// TIA Portal V19 export
DATA_BLOCK "CV_DATA"   // DB17
{ S7_Optimized_Access := 'FALSE' }
   VAR
      CHILLED_SKID_P01 : Struct
         CMD : Bool;
         SET_POINT : Real;
         INPUT : Real;
         OUT_PUT : Real;
         OUTPUT_PER : Int;
         NORM_MIN : Int;
         NORM_MAX : Int := 27684;
         NORM_OUT : Real;
         SCALE_MIN : Real;
         SCALE_MAX : Real := 50.0;
         SCALE_OUT : Real;
         MANUAL_OPEN_PER : Int;
         MANUAL_TEMP : Int;
         MANOUT : Real;
         PUMP_AO : Real;
      END_STRUCT;
      HS_PCV801 : Struct
         CMD : Bool;
         SET_POINT : Real;
         INPUT : Real;
         OUT_PUT : Real;
         OUTPUT_PER : Int;
         NORM_MIN : Int;
         NORM_MAX : Int;
         NORM_OUT : Real;
         SCALE_MIN : Real;
         SCALE_MAX : Real;
         SCALE_OUT : Real;
         MANUAL_OPEN_PER : Int;
         MANUAL_TEMP : Int;
         MANOUT : Int;
         CV_AO : Int;
      END_STRUCT;
      CHILLED_SKID_P02 : Struct
         CMD : Bool;
         SET_POINT : Real;
         INPUT : Real;
         OUT_PUT : Real;
         OUTPUT_PER : Int;
         NORM_MIN : Int;
         NORM_MAX : Int := 27684;
         NORM_OUT : Real := 0.0;
         SCALE_MIN : Real := 0.0;
         SCALE_MAX : Real := 50.0;
         SCALE_OUT : Real;
         MANUAL_OPEN_PER : Int;
         MANUAL_TEMP : Int;
         MANOUT : Real;
         PUMP_AO : Real;
      END_STRUCT;
      CHILLED_SKID_P03 : Struct
         CMD : Bool;
         SET_POINT : Real;
         INPUT : Real;
         OUT_PUT : Real;
         OUTPUT_PER : Int;
         NORM_MIN : Int;
         NORM_MAX : Int := 27684;
         NORM_OUT : Real := 0.0;
         SCALE_MIN : Real := 0.0;
         SCALE_MAX : Real := 50.0;
         SCALE_OUT : Real;
         MANUAL_OPEN_PER : Int;
         MANUAL_TEMP : Int;
         MANOUT : Real;
         PUMP_AO : Real;
      END_STRUCT;
      HOT_SKID_P01 : Struct
         CMD : Bool;
         SET_POINT : Real;
         INPUT : Real;
         OUT_PUT : Real;
         OUTPUT_PER : Int;
         NORM_MIN : Int;
         NORM_MAX : Int := 27684;
         NORM_OUT : Real := 0.0;
         SCALE_MIN : Real := 0.0;
         SCALE_MAX : Real := 50.0;
         SCALE_OUT : Real;
         MANUAL_OPEN_PER : Int;
         MANUAL_TEMP : Int;
         MANOUT : Real;
         PUMP_AO : Real;
      END_STRUCT;
      HOT_SKID_P02 : Struct
         CMD : Bool;
         SET_POINT : Real;
         INPUT : Real;
         OUT_PUT : Real;
         OUTPUT_PER : Int;
         NORM_MIN : Int;
         NORM_MAX : Int := 27684;
         NORM_OUT : Real := 0.0;
         SCALE_MIN : Real := 0.0;
         SCALE_MAX : Real := 50.0;
         SCALE_OUT : Real;
         MANUAL_OPEN_PER : Int;
         MANUAL_TEMP : Int;
         MANOUT : Real;
         PUMP_AO : Real;
      END_STRUCT;
      HOT_SKID_P03 : Struct
         CMD : Bool;
         SET_POINT : Real;
         INPUT : Real;
         OUT_PUT : Real;
         OUTPUT_PER : Int;
         NORM_MIN : Int;
         NORM_MAX : Int := 27684;
         NORM_OUT : Real := 0.0;
         SCALE_MIN : Real := 0.0;
         SCALE_MAX : Real := 50.0;
         SCALE_OUT : Real;
         MANUAL_OPEN_PER : Int;
         MANUAL_TEMP : Int;
         MANOUT : Real;
         PUMP_AO : Real;
      END_STRUCT;
      COLD_SKID_P01 : Struct
         CMD : Bool;
         SET_POINT : Real;
         INPUT : Real;
         OUT_PUT : Real;
         OUTPUT_PER : Int;
         NORM_MIN : Int;
         NORM_MAX : Int := 27684;
         NORM_OUT : Real := 0.0;
         SCALE_MIN : Real := 0.0;
         SCALE_MAX : Real := 50.0;
         SCALE_OUT : Real;
         MANUAL_OPEN_PER : Int;
         MANUAL_TEMP : Int;
         MANOUT : Real;
         PUMP_AO : Real;
      END_STRUCT;
      COLD_SKID_P02 : Struct
         CMD : Bool;
         SET_POINT : Real;
         INPUT : Real;
         OUT_PUT : Real;
         OUTPUT_PER : Int;
         NORM_MIN : Int;
         NORM_MAX : Int := 27684;
         NORM_OUT : Real := 0.0;
         SCALE_MIN : Real := 0.0;
         SCALE_MAX : Real := 50.0;
         SCALE_OUT : Real;
         MANUAL_OPEN_PER : Int;
         MANUAL_TEMP : Int;
         MANOUT : Real;
         PUMP_AO : Real;
      END_STRUCT;
      COLD_SKID_P03 : Struct
         CMD : Bool;
         SET_POINT : Real;
         INPUT : Real;
         OUT_PUT : Real;
         OUTPUT_PER : Int;
         NORM_MIN : Int;
         NORM_MAX : Int := 27684;
         NORM_OUT : Real := 0.0;
         SCALE_MIN : Real := 0.0;
         SCALE_MAX : Real := 50.0;
         SCALE_OUT : Real;
         MANUAL_OPEN_PER : Int;
         MANUAL_TEMP : Int;
         MANOUT : Real;
         PUMP_AO : Real;
      END_STRUCT;
      UCH_SKID_P01 : Struct
         CMD : Bool;
         SET_POINT : Real;
         INPUT : Real;
         OUT_PUT : Real;
         OUTPUT_PER : Int;
         NORM_MIN : Int;
         NORM_MAX : Int := 27684;
         NORM_OUT : Real := 0.0;
         SCALE_MIN : Real := 0.0;
         SCALE_MAX : Real := 50.0;
         SCALE_OUT : Real;
         MANUAL_OPEN_PER : Int;
         MANUAL_TEMP : Int;
         MANOUT : Real;
         PUMP_AO : Real;
      END_STRUCT;
      UCH_SKID_P02 : Struct
         CMD : Bool;
         SET_POINT : Real;
         INPUT : Real;
         OUT_PUT : Real;
         OUTPUT_PER : Int;
         NORM_MIN : Int;
         NORM_MAX : Int := 27684;
         NORM_OUT : Real := 0.0;
         SCALE_MIN : Real := 0.0;
         SCALE_MAX : Real := 50.0;
         SCALE_OUT : Real;
         MANUAL_OPEN_PER : Int;
         MANUAL_TEMP : Int;
         MANOUT : Real;
         PUMP_AO : Real;
      END_STRUCT;
   END_VAR
BEGIN
END_DATA_BLOCK
